// TIA Portal V21 export
// export: Created 2026-10-23T20:44:41.5268196Z, ExportSetting WithDefaults, DisplayName Totally Integrated Automation Portal, DisplayVersion V21 Update 1, DisplayName SINAMICS Startdrive Advanced, DisplayVersion V21 HF2, DisplayName SINAMICS Startdrive G110M, G120, G120C, G120D, G120P, G115D, DisplayVersion V21 HF2, DisplayName SINAMICS Startdrive G130, G150, S120, S150, G200, G220, S200, S210, S220, Innomotics MVD, DisplayVersion V21 HF2, DisplayName STEP 7 Professional, DisplayVersion V21 Update 1, DisplayName STEP 7 Safety, DisplayVersion V21, DisplayName Tech WebApplication, DisplayVersion V21, DisplayName WinCC Basic/Comfort/Advanced, DisplayVersion V21 Update 1, DisplayName WinCC Unified, DisplayVersion V21 Update 1
ORGANIZATION_BLOCK "OB_Dosing"   // OB124, SCL, ProgramCycle
TITLE = "Main Program Sweep (Cycle)" / Dosing cycle
VERSION : 0.1
// Program cycle OB of the unit Dosing; calls FB_Doser
// stored: AutoNumber true, IsIECCheckEnabled false, Namespace Dosing, SetENOAutomatically false
   VAR_INPUT
      Initial_Call : Bool;   // Initial call of this OB
      Remanence : Bool;   // =True, if remanent data are available
   END_VAR
BEGIN

       "Dosing.IDB_Doser"(Start := TRUE, Stop := FALSE);
END_ORGANIZATION_BLOCK
